// TIA Portal V21 export
GraphicList "GL_BitNo"  ListRange=Binary
  GraphicListEntry   EntryType=SingleValue, Picture=G_PNG
  GraphicListEntry   EntryType=SingleValue, From=1, To=1, Picture=G_JPG
  GraphicListEntry   EntryType=SingleValue, From=2, To=2, Picture=G_BMP
  GraphicListEntry   EntryType=SingleValue, From=3, To=3, Picture=G_TIF
